TYPE "ST_SignalTowerParCfg"
VERSION : 0.1
   STRUCT
      SchemaVersion : UInt := 1;
      LampTestDuration : Time := T#3S;
      OperatorUsesWhite : Bool;
      HornOnHigh : Bool := TRUE;
   END_STRUCT;

END_TYPE

